{attribute 'Tc2GvlVarNames'}
VAR_GLOBAL CONSTANT
	nZONES_MAX_NO			:UINT := 4;			(* Amount of control zones *)
END_VAR

(* stored: Version 1.1.0.1, ProductVersion 3.1.4024.15
   GVL GVL_FB_GFX4IRZones: Id {e5446c59-c3d5-4e2f-b326-9c3b97416d8d} *)
